(* PLC project fbd_reactor_2oo3_clean, Anonymous Benchmark Suite 1.0 *)
(* stored: creationDateTime 2026-08-26T00:00:00 *)

PROGRAM trip_logic
  VAR_INPUT
    ps1 : BOOL;
    ps2 : BOOL;
    ps3 : BOOL;
  END_VAR
  VAR_OUTPUT
    trip : BOOL;
  END_VAR

(* FBD diagram, written out as Structured Text *)
trip := ps1 AND ps2 OR ps2 AND ps3 OR ps1 AND ps3;
END_PROGRAM

CONFIGURATION Config0
  RESOURCE Res0 ON PLC
    TASK tcyclic(INTERVAL := T#10ms, PRIORITY := 0);
    PROGRAM inst0 WITH tcyclic : trip_logic;
  END_RESOURCE
END_CONFIGURATION
